// TIA Portal V20 export
DATA_BLOCK "Verwaltung_Teiledaten_FB_DB"   // DB1
// stored: InstanceOfName Verwaltung_Teiledaten_FB, InstanceOfType FB
"Verwaltung_Teiledaten_FB"
BEGIN
END_DATA_BLOCK
